(* Logix 5000 project; controller TFF vendor 1 type 14 code 107 rev 33.11; software revision 33.04; part 26 of 38 *)
(* tags used below, declared in another part *)
   Address : DINT;   // Temp Address
   Index : DINT;   // Index
   PCV101_PID_Settings : INT;
   TIME : DINT[2];
   AnalogOutput : AnalogOutput[25];   // Analog Output Array
   AnalogPoint : AnalogInput[50];   // Analog Input Array
   ControlLoop : ControlLoop[20];   // Control Loop Array
   ControlLoop_PCV201 : ALIAS FOR ControlLoop[5];
   ControlLoop_PCV201_5ms : ALIAS FOR ControlLoop[6];
   ControlLoop_PCV201_CV : REAL;   // Control Value
   ControlLoop_PCV201_RAMP_OUT : REAL;   // Ramp Output
   ControlLoop_TIC101 : ALIAS FOR ControlLoop[7];
   ExternalTCU : BOOL;   // Use of External TCU
   LI101 : ALIAS FOR AnalogPoint[44];
   PCV201_Control : PCV_Control;   // PCV201 Control UDT
   Phase0 : ALIAS FOR Phase[0];   // Phase 0
   SysControl : SysControl;   // General system status and command
   Tank : TankManagement;   // Tank Management
   TCU101_AO : ALIAS FOR AnalogOutput[6];
   TCU101ON : ALIAS FOR DigitalOutput[20];
   TIC101Control : TCUControl;
(* Process, continued *)

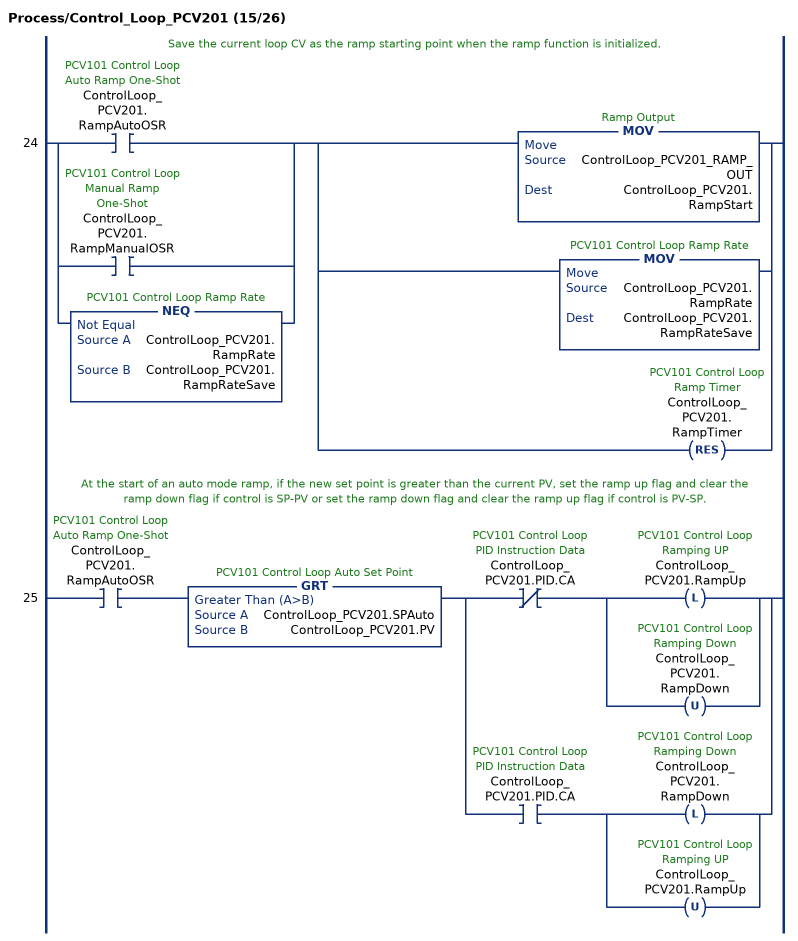
   [picture p239: Process/Control_Loop_PCV201 rungs 24-25]
   // Save the current loop CV as the ramp starting point when the ramp function is initialized.
   24: [XIC(ControlLoop_PCV201.RampAutoOSR) ,XIC(ControlLoop_PCV201.RampManualOSR) ,NEQ(ControlLoop_PCV201.RampRate,ControlLoop_PCV201.RampRateSave) ][MOV(ControlLoop_PCV201_RAMP_OUT,ControlLoop_PCV201.RampStart) ,MOV(ControlLoop_PCV201.RampRate,ControlLoop_PCV201.RampRateSave) ,RES(ControlLoop_PCV201.RampTimer) ];
   // At the start of an auto mode ramp, if the new set point is greater than the current PV, set the ramp up flag and clear the ramp down flag if control is SP-PV or set the ramp down flag and clear the ramp up flag if control is PV-SP.
   25: XIC(ControlLoop_PCV201.RampAutoOSR)GRT(ControlLoop_PCV201.SPAuto,ControlLoop_PCV201.PV)[XIO(ControlLoop_PCV201.PID.CA) [OTL(ControlLoop_PCV201.RampUp) ,OTU(ControlLoop_PCV201.RampDown) ] ,XIC(ControlLoop_PCV201.PID.CA) [OTL(ControlLoop_PCV201.RampDown) ,OTU(ControlLoop_PCV201.RampUp) ] ];
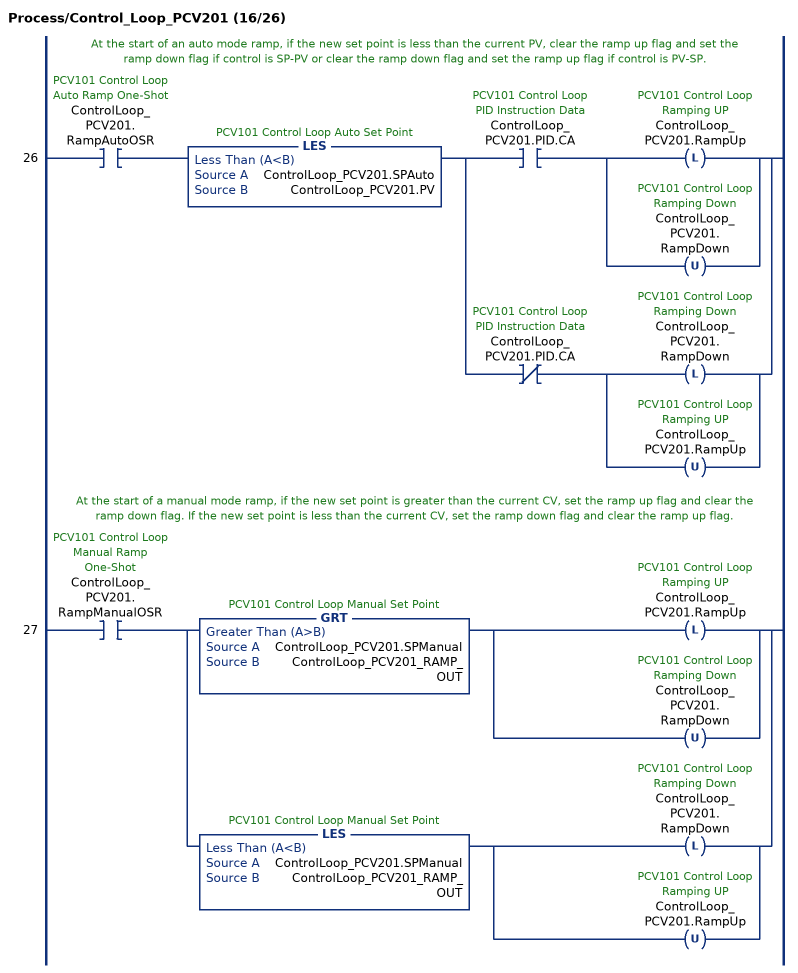
   // At the start of an auto mode ramp, if the new set point is less than the current PV, clear the ramp up flag and set the ramp down flag if control is SP-PV or clear the ramp down flag and set the ramp up flag if control is PV-SP.
   26: XIC(ControlLoop_PCV201.RampAutoOSR)LES(ControlLoop_PCV201.SPAuto,ControlLoop_PCV201.PV)[XIC(ControlLoop_PCV201.PID.CA) [OTL(ControlLoop_PCV201.RampUp) ,OTU(ControlLoop_PCV201.RampDown) ] ,XIO(ControlLoop_PCV201.PID.CA) [OTL(ControlLoop_PCV201.RampDown) ,OTU(ControlLoop_PCV201.RampUp) ] ];
   // At the start of a manual mode ramp, if the new set point is greater than the current CV, set the ramp up flag and clear the ramp down flag. If the new set point is less than the current CV, set the ramp down flag and clear the ramp up flag.
   27: XIC(ControlLoop_PCV201.RampManualOSR)[GRT(ControlLoop_PCV201.SPManual,ControlLoop_PCV201_RAMP_OUT) [OTL(ControlLoop_PCV201.RampUp) ,OTU(ControlLoop_PCV201.RampDown) ] ,LES(ControlLoop_PCV201.SPManual,ControlLoop_PCV201_RAMP_OUT) [OTL(ControlLoop_PCV201.RampDown) ,OTU(ControlLoop_PCV201.RampUp) ] ];
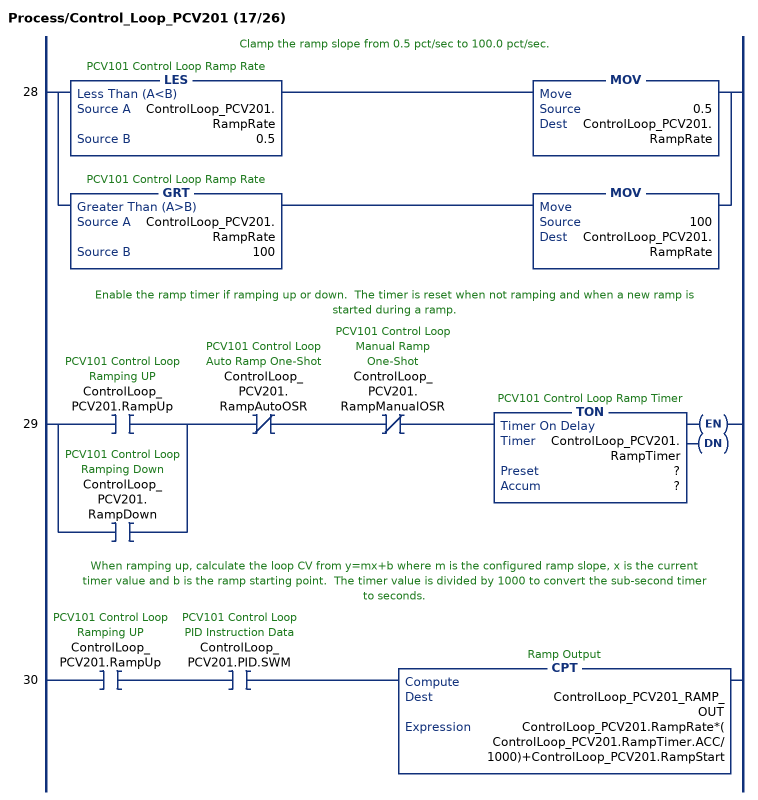
   // Clamp the ramp slope from 0.5 pct/sec to 100.0 pct/sec.
   28: [LES(ControlLoop_PCV201.RampRate,0.5) MOV(0.5,ControlLoop_PCV201.RampRate) ,GRT(ControlLoop_PCV201.RampRate,100) MOV(100,ControlLoop_PCV201.RampRate) ];
   // Enable the ramp timer if ramping up or down.  The timer is reset when not ramping and when a new ramp is started during a ramp.
   29: [XIC(ControlLoop_PCV201.RampUp) ,XIC(ControlLoop_PCV201.RampDown) ]XIO(ControlLoop_PCV201.RampAutoOSR)XIO(ControlLoop_PCV201.RampManualOSR)TON(ControlLoop_PCV201.RampTimer,?,?);
   // When ramping up, calculate the loop CV from y=mx+b where m is the configured ramp slope, x is the current timer value and b is the ramp starting point.  The timer value is divided by 1000 to convert the sub-second timer to seconds.
   30: XIC(ControlLoop_PCV201.RampUp)XIC(ControlLoop_PCV201.PID.SWM)CPT(ControlLoop_PCV201_RAMP_OUT,ControlLoop_PCV201.RampRate*(ControlLoop_PCV201.RampTimer.ACC/1000)+ControlLoop_PCV201.RampStart);
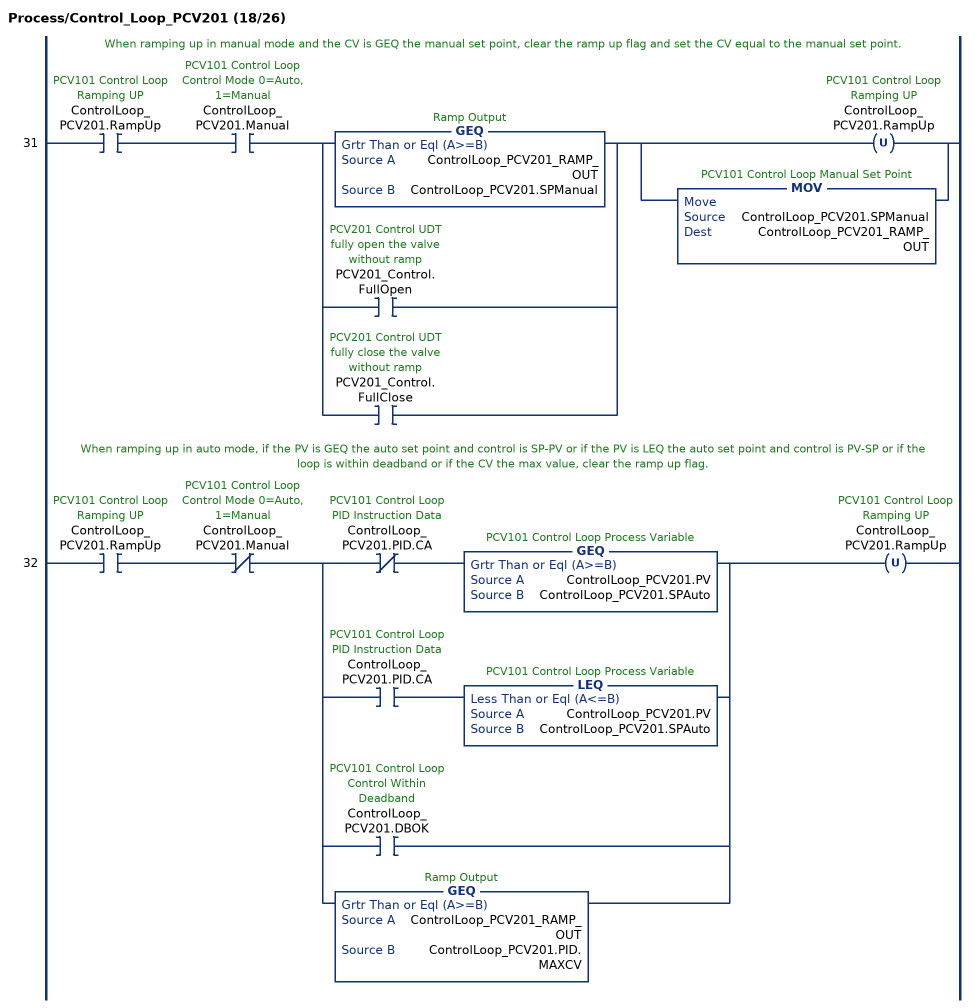
   // When ramping up in manual mode and the CV is GEQ the manual set point, clear the ramp up flag and set the CV equal to the manual set point.
   31: XIC(ControlLoop_PCV201.RampUp)XIC(ControlLoop_PCV201.Manual)[GEQ(ControlLoop_PCV201_RAMP_OUT,ControlLoop_PCV201.SPManual) ,XIC(PCV201_Control.FullOpen) ,XIC(PCV201_Control.FullClose) ][OTU(ControlLoop_PCV201.RampUp) ,MOV(ControlLoop_PCV201.SPManual,ControlLoop_PCV201_RAMP_OUT) ];
   // When ramping up in auto mode, if the PV is GEQ the auto set point and control is SP-PV or if the PV is LEQ the auto set point and control is PV-SP or if the loop is within deadband or if the CV the max value, clear the ramp up flag.
   32: XIC(ControlLoop_PCV201.RampUp)XIO(ControlLoop_PCV201.Manual)[XIO(ControlLoop_PCV201.PID.CA) GEQ(ControlLoop_PCV201.PV,ControlLoop_PCV201.SPAuto) ,XIC(ControlLoop_PCV201.PID.CA) LEQ(ControlLoop_PCV201.PV,ControlLoop_PCV201.SPAuto) ,XIC(ControlLoop_PCV201.DBOK) ,GEQ(ControlLoop_PCV201_RAMP_OUT,ControlLoop_PCV201.PID.MAXCV) ]OTU(ControlLoop_PCV201.RampUp);
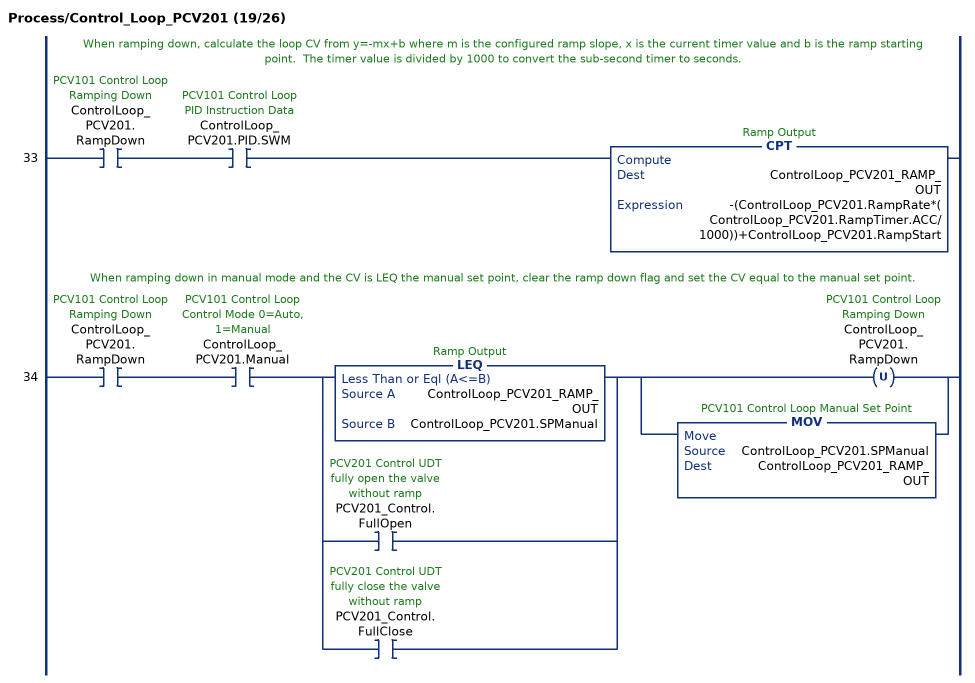
   // When ramping down, calculate the loop CV from y=-mx+b where m is the configured ramp slope, x is the current timer value and b is the ramp starting point.  The timer value is divided by 1000 to convert the sub-second timer to seconds.
   33: XIC(ControlLoop_PCV201.RampDown)XIC(ControlLoop_PCV201.PID.SWM)CPT(ControlLoop_PCV201_RAMP_OUT,-(ControlLoop_PCV201.RampRate*(ControlLoop_PCV201.RampTimer.ACC/1000))+ControlLoop_PCV201.RampStart);
   // When ramping down in manual mode and the CV is LEQ the manual set point, clear the ramp down flag and set the CV equal to the manual set point.
   34: XIC(ControlLoop_PCV201.RampDown)XIC(ControlLoop_PCV201.Manual)[LEQ(ControlLoop_PCV201_RAMP_OUT,ControlLoop_PCV201.SPManual) ,XIC(PCV201_Control.FullOpen) ,XIC(PCV201_Control.FullClose) ][OTU(ControlLoop_PCV201.RampDown) ,MOV(ControlLoop_PCV201.SPManual,ControlLoop_PCV201_RAMP_OUT) ];
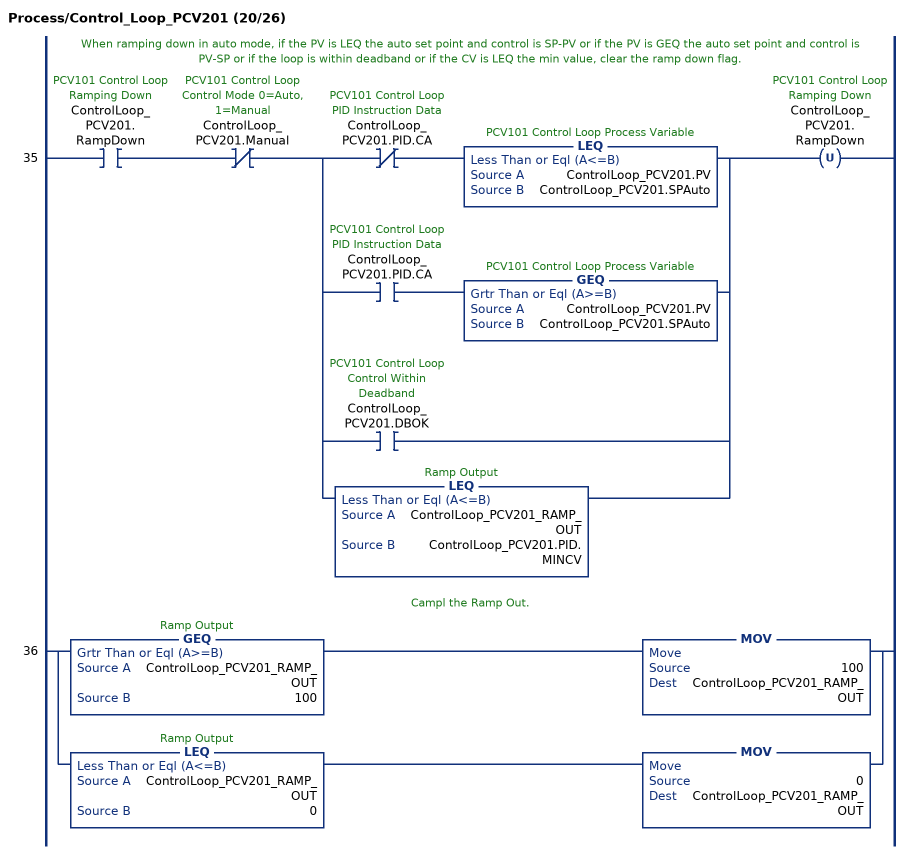
   // When ramping down in auto mode, if the PV is LEQ the auto set point and control is SP-PV or if the PV is GEQ the auto set point and control is PV-SP or if the loop is within deadband or if the CV is LEQ the min value, clear the ramp down flag.
   35: XIC(ControlLoop_PCV201.RampDown)XIO(ControlLoop_PCV201.Manual)[XIO(ControlLoop_PCV201.PID.CA) LEQ(ControlLoop_PCV201.PV,ControlLoop_PCV201.SPAuto) ,XIC(ControlLoop_PCV201.PID.CA) GEQ(ControlLoop_PCV201.PV,ControlLoop_PCV201.SPAuto) ,XIC(ControlLoop_PCV201.DBOK) ,LEQ(ControlLoop_PCV201_RAMP_OUT,ControlLoop_PCV201.PID.MINCV) ]OTU(ControlLoop_PCV201.RampDown);
   // Campl the Ramp Out.
   36: [GEQ(ControlLoop_PCV201_RAMP_OUT,100) MOV(100,ControlLoop_PCV201_RAMP_OUT) ,LEQ(ControlLoop_PCV201_RAMP_OUT,0) MOV(0,ControlLoop_PCV201_RAMP_OUT) ];
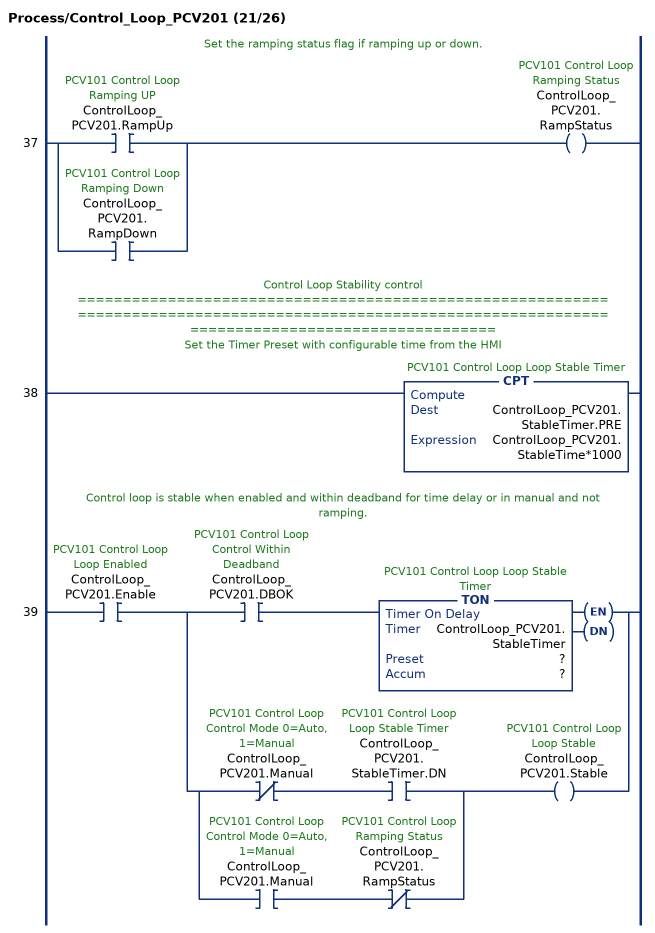
   // Set the ramping status flag if ramping up or down.
   37: [XIC(ControlLoop_PCV201.RampUp) ,XIC(ControlLoop_PCV201.RampDown) ]OTE(ControlLoop_PCV201.RampStatus);
   // Control Loop Stability control
   // ========================================================================================================================================================
   // Set the Timer Preset with configurable time from the HMI
   38: CPT(ControlLoop_PCV201.StableTimer.PRE,ControlLoop_PCV201.StableTime*1000);
   // Control loop is stable when enabled and within deadband for time delay or in manual and not ramping.
   39: XIC(ControlLoop_PCV201.Enable)[XIC(ControlLoop_PCV201.DBOK) TON(ControlLoop_PCV201.StableTimer,?,?) ,[XIO(ControlLoop_PCV201.Manual) XIC(ControlLoop_PCV201.StableTimer.DN) ,XIC(ControlLoop_PCV201.Manual) XIO(ControlLoop_PCV201.RampStatus) ] OTE(ControlLoop_PCV201.Stable) ];
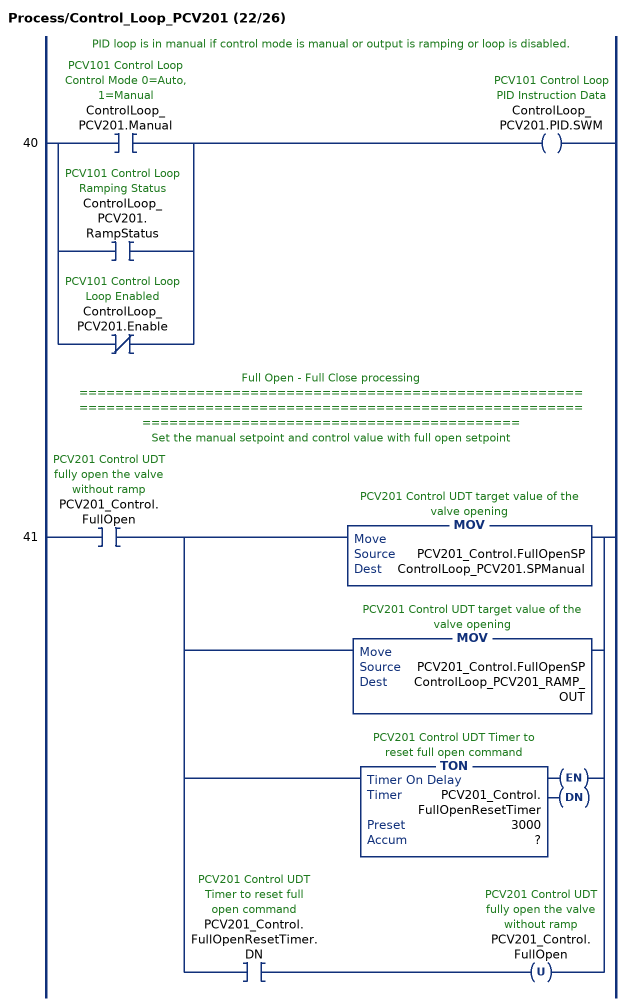
   // PID loop is in manual if control mode is manual or output is ramping or loop is disabled.
   40: [XIC(ControlLoop_PCV201.Manual) ,XIC(ControlLoop_PCV201.RampStatus) ,XIO(ControlLoop_PCV201.Enable) ]OTE(ControlLoop_PCV201.PID.SWM);
   // Full Open - Full Close processing
   // ==========================================================================================================================================================
   // Set the manual setpoint and control value with full open setpoint
   41: XIC(PCV201_Control.FullOpen)[MOV(PCV201_Control.FullOpenSP,ControlLoop_PCV201.SPManual) ,MOV(PCV201_Control.FullOpenSP,ControlLoop_PCV201_RAMP_OUT) ,TON(PCV201_Control.FullOpenResetTimer,?,?) ,XIC(PCV201_Control.FullOpenResetTimer.DN) OTU(PCV201_Control.FullOpen) ];
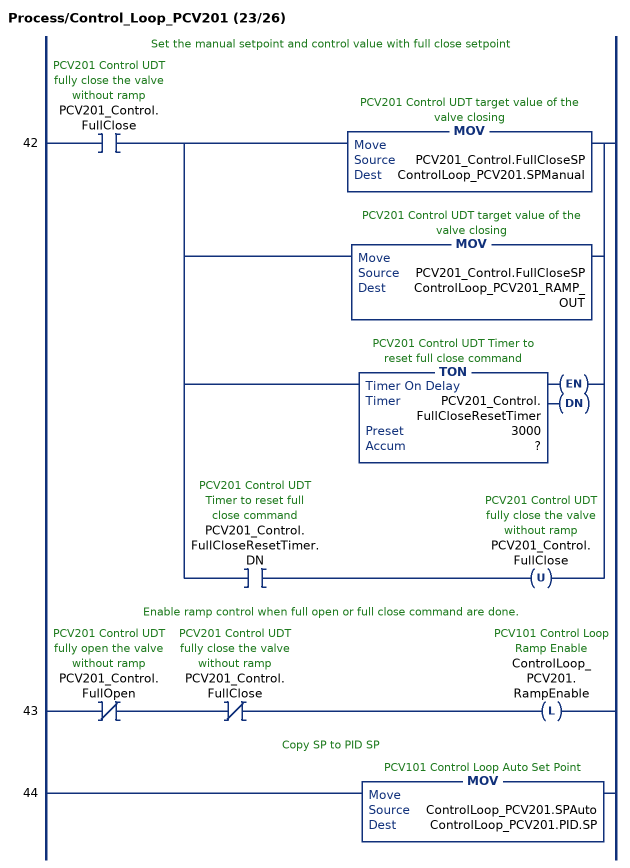
   // Set the manual setpoint and control value with full close setpoint
   42: XIC(PCV201_Control.FullClose)[MOV(PCV201_Control.FullCloseSP,ControlLoop_PCV201.SPManual) ,MOV(PCV201_Control.FullCloseSP,ControlLoop_PCV201_RAMP_OUT) ,TON(PCV201_Control.FullCloseResetTimer,?,?) ,XIC(PCV201_Control.FullCloseResetTimer.DN) OTU(PCV201_Control.FullClose) ];
   // Enable ramp control when full open or full close command are done.
   43: XIO(PCV201_Control.FullOpen)XIO(PCV201_Control.FullClose)OTL(ControlLoop_PCV201.RampEnable);
   // Copy SP to PID SP
   44: MOV(ControlLoop_PCV201.SPAuto,ControlLoop_PCV201.PID.SP);
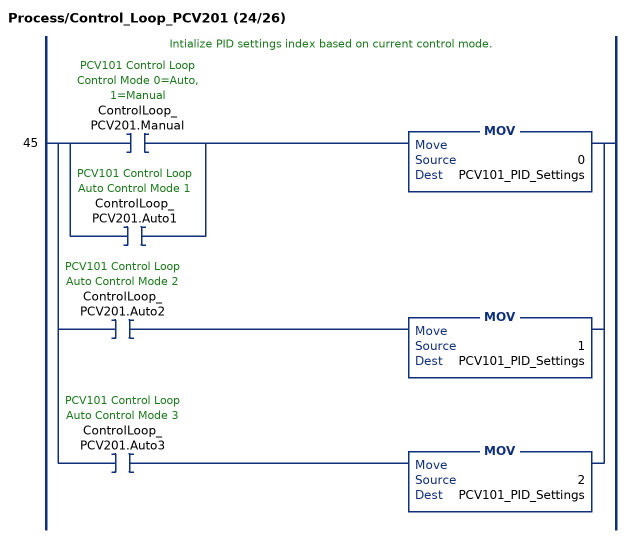
   // Intialize PID settings index based on current control mode.
   45: [[XIC(ControlLoop_PCV201.Manual) ,XIC(ControlLoop_PCV201.Auto1) ] MOV(0,PCV101_PID_Settings) ,XIC(ControlLoop_PCV201.Auto2) MOV(1,PCV101_PID_Settings) ,XIC(ControlLoop_PCV201.Auto3) MOV(2,PCV101_PID_Settings) ];
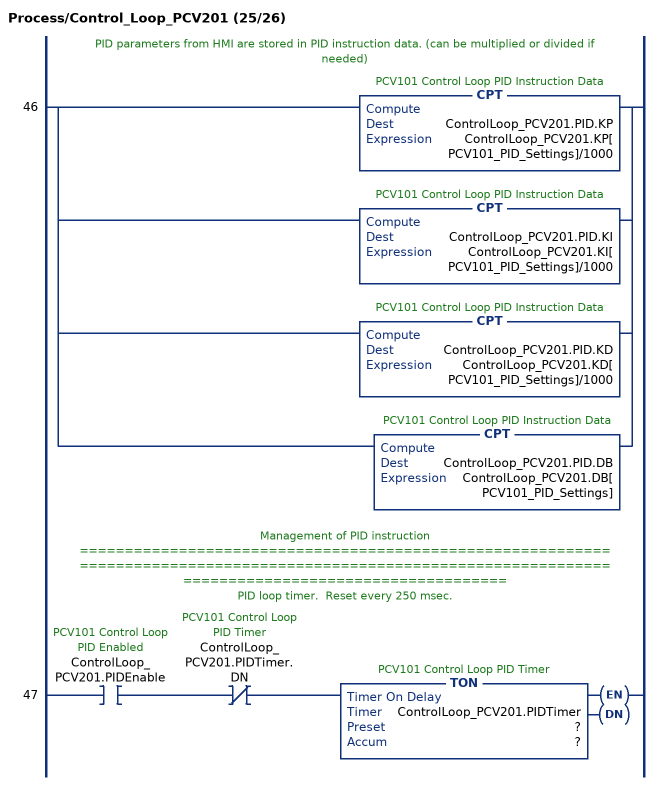
   // PID parameters from HMI are stored in PID instruction data. (can be multiplied or divided if needed)
   46: [CPT(ControlLoop_PCV201.PID.KP,ControlLoop_PCV201.KP[PCV101_PID_Settings]/1000) ,CPT(ControlLoop_PCV201.PID.KI,ControlLoop_PCV201.KI[PCV101_PID_Settings]/1000) ,CPT(ControlLoop_PCV201.PID.KD,ControlLoop_PCV201.KD[PCV101_PID_Settings]/1000) ,CPT(ControlLoop_PCV201.PID.DB,ControlLoop_PCV201.DB[PCV101_PID_Settings]) ];
   // Management of PID instruction
   // ==========================================================================================================================================================
   // PID loop timer.  Reset every 250 msec.
   47: XIC(ControlLoop_PCV201.PIDEnable)XIO(ControlLoop_PCV201.PIDTimer.DN)TON(ControlLoop_PCV201.PIDTimer,?,?);
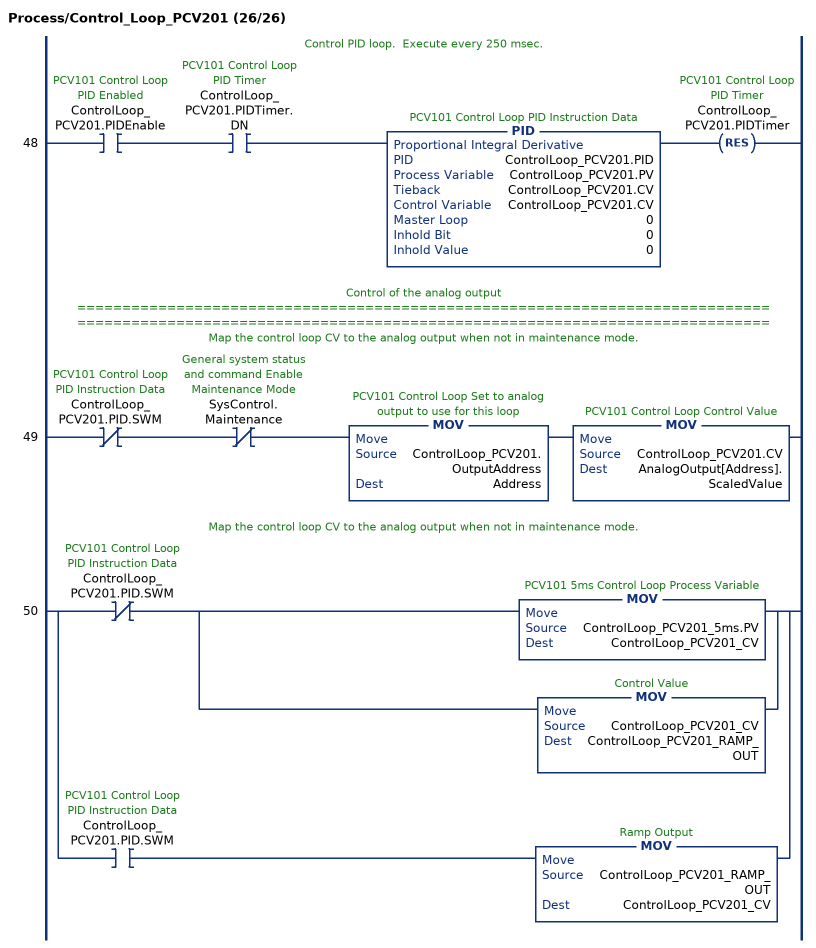
   // Control PID loop.  Execute every 250 msec.
   48: XIC(ControlLoop_PCV201.PIDEnable)XIC(ControlLoop_PCV201.PIDTimer.DN)PID(ControlLoop_PCV201.PID,ControlLoop_PCV201.PV,ControlLoop_PCV201.CV,ControlLoop_PCV201.CV,0,0,0)RES(ControlLoop_PCV201.PIDTimer);
   // Control of the analog output
   // ==========================================================================================================================================================
   // Map the control loop CV to the analog output when not in maintenance mode.
   49: XIO(ControlLoop_PCV201.PID.SWM)XIO(SysControl.Maintenance)MOV(ControlLoop_PCV201.OutputAddress,Address)MOV(ControlLoop_PCV201.CV,AnalogOutput[Address].ScaledValue);
   // Map the control loop CV to the analog output when not in maintenance mode.
   50: [XIO(ControlLoop_PCV201.PID.SWM) [MOV(ControlLoop_PCV201_5ms.PV,ControlLoop_PCV201_CV) ,MOV(ControlLoop_PCV201_CV,ControlLoop_PCV201_RAMP_OUT) ] ,XIC(ControlLoop_PCV201.PID.SWM) MOV(ControlLoop_PCV201_RAMP_OUT,ControlLoop_PCV201_CV) ];
END_ROUTINE

ROUTINE Control_Loop_TIC101   (* ladder *)
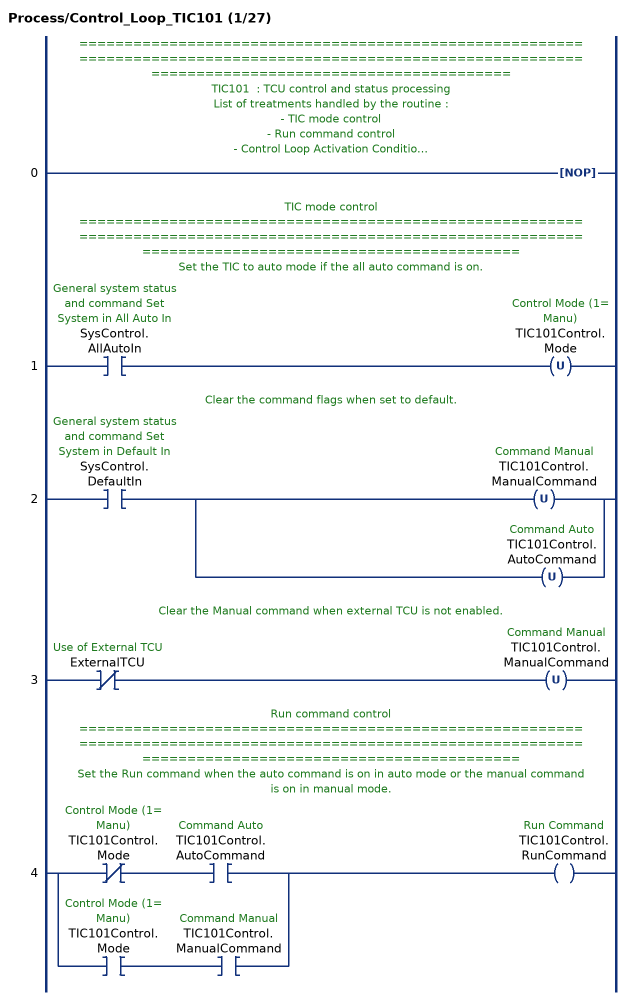
   // ========================================================================================================================================================
   //                                                                                                    TIC101  : TCU control and status processing
   //                                                     List of treatments handled by the routine :
   //                                                     - TIC mode control
   //                                                        - Run command control
   //                                                          - Control Loop Activation Condition
   //                                                          - Control Loop initialization
   //                                                          - Mode control
   //                                                          - Control Loop deadband calculation
   //                                                          - Management of ramping control
   //                                                            - Management of SP Offset
   //                                                          - Control Loop Stability control
   //                                                          - Control Loop manual state control
   //                                                          - Management of PID instruction
   //                                                          - Control of the analog output
   //                                                     -----------------------------------------------------------------------------------------------------------------------------------------------------
   //                                                     History
   // 		2019-DEC-24 - Merck - Q. Spindler - Initial version for Candidate Release 1.00.00.00.a
   // 		2020-SEP-09 - Merck - Q. Spindler - Modifications for Candidate Release 1.00.00.00.d
   // 					- Add ControlLoop Enable and not manual condition for DBOK status
   // 				   	- Clear Manual command when ExternalTCU is disabled
   // 		2021-APR-16 - Merck - Q. Spindler - Modifications for Candidate Release 1.00.00.00.e
   //                                        - Add Initialize address if no mode selected.
   //                       - Change TIC Output Range to 50
   // ========================================================================================================================================================
   0: NOP();
   // TIC mode control
   // ==========================================================================================================================================================
   // Set the TIC to auto mode if the all auto command is on.
   1: XIC(SysControl.AllAutoIn)OTU(TIC101Control.Mode);
   // Clear the command flags when set to default.
   2: XIC(SysControl.DefaultIn)[OTU(TIC101Control.ManualCommand) ,OTU(TIC101Control.AutoCommand) ];
   // Clear the Manual command when external TCU is not enabled.
   3: XIO(ExternalTCU)OTU(TIC101Control.ManualCommand);
   // Run command control
   // ==========================================================================================================================================================
   // Set the Run command when the auto command is on in auto mode or the manual command is on in manual mode.
   4: [XIO(TIC101Control.Mode) XIC(TIC101Control.AutoCommand) ,XIC(TIC101Control.Mode) XIC(TIC101Control.ManualCommand) ]OTE(TIC101Control.RunCommand);
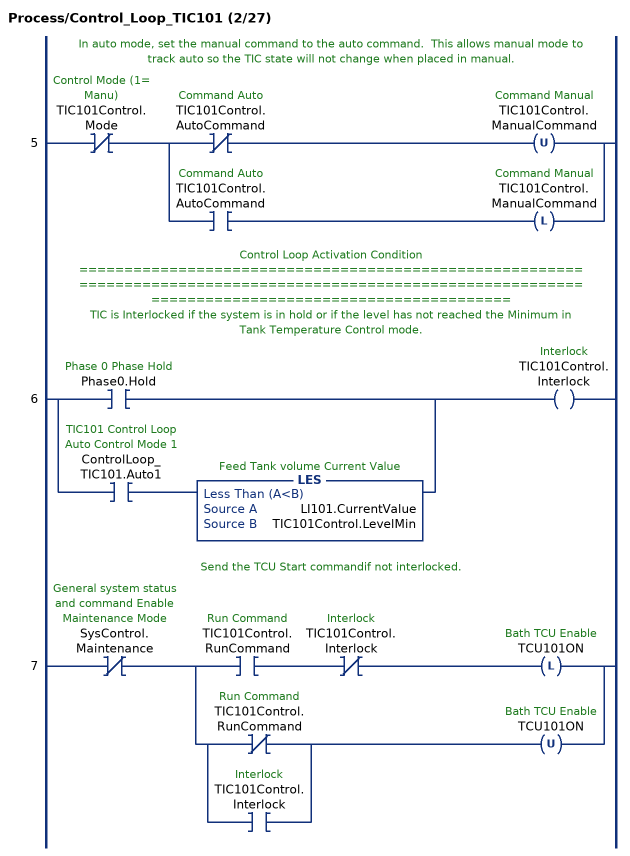
   // In auto mode, set the manual command to the auto command.  This allows manual mode to track auto so the TIC state will not change when placed in manual.
   5: XIO(TIC101Control.Mode)[XIO(TIC101Control.AutoCommand) OTU(TIC101Control.ManualCommand) ,XIC(TIC101Control.AutoCommand) OTL(TIC101Control.ManualCommand) ];
   // Control Loop Activation Condition
   // ========================================================================================================================================================
   // TIC is Interlocked if the system is in hold or if the level has not reached the Minimum in Tank Temperature Control mode.
   6: [XIC(Phase0.Hold) ,XIC(ControlLoop_TIC101.Auto1) LES(LI101.CurrentValue,TIC101Control.LevelMin) ]OTE(TIC101Control.Interlock);
   // Send the TCU Start commandif not interlocked.
   7: XIO(SysControl.Maintenance)[XIC(TIC101Control.RunCommand) XIO(TIC101Control.Interlock) OTL(TCU101ON) ,[XIO(TIC101Control.RunCommand) ,XIC(TIC101Control.Interlock) ] OTU(TCU101ON) ];
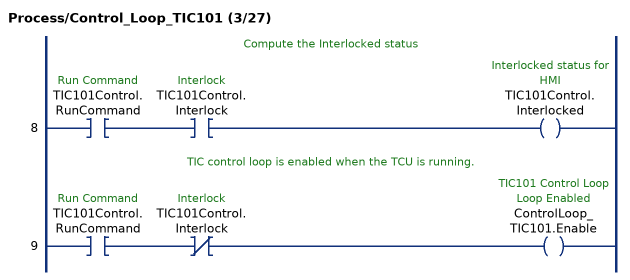
   // Compute the Interlocked status
   8: XIC(TIC101Control.RunCommand)XIC(TIC101Control.Interlock)OTE(TIC101Control.Interlocked);
   // TIC control loop is enabled when the TCU is running.
   9: XIC(TIC101Control.RunCommand)XIO(TIC101Control.Interlock)OTE(ControlLoop_TIC101.Enable);
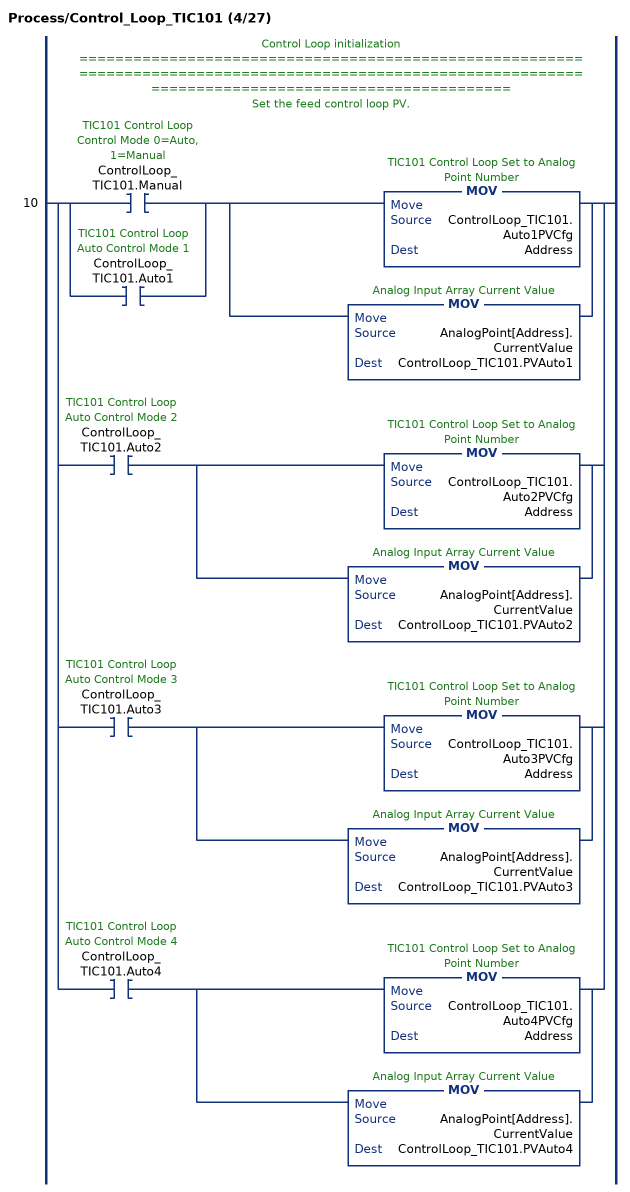
   // Control Loop initialization
   // ========================================================================================================================================================
   // Set the feed control loop PV.
   10: [[[XIC(ControlLoop_TIC101.Manual) ,XIC(ControlLoop_TIC101.Auto1) ] [MOV(ControlLoop_TIC101.Auto1PVCfg,Address) ,MOV(AnalogPoint[Address].CurrentValue,ControlLoop_TIC101.PVAuto1) ] ,XIC(ControlLoop_TIC101.Auto2) [MOV(ControlLoop_TIC101.Auto2PVCfg,Address) ,MOV(AnalogPoint[Address].CurrentValue,ControlLoop_TIC101.PVAuto2) ] ] ,XIC(ControlLoop_TIC101.Auto3) [MOV(ControlLoop_TIC101.Auto3PVCfg,Address) ,MOV(AnalogPoint[Address].CurrentValue,ControlLoop_TIC101.PVAuto3) ] ,XIC(ControlLoop_TIC101.Auto4) [MOV(ControlLoop_TIC101.Auto4PVCfg,Address) ,MOV(AnalogPoint[Address].CurrentValue,ControlLoop_TIC101.PVAuto4) ] ];
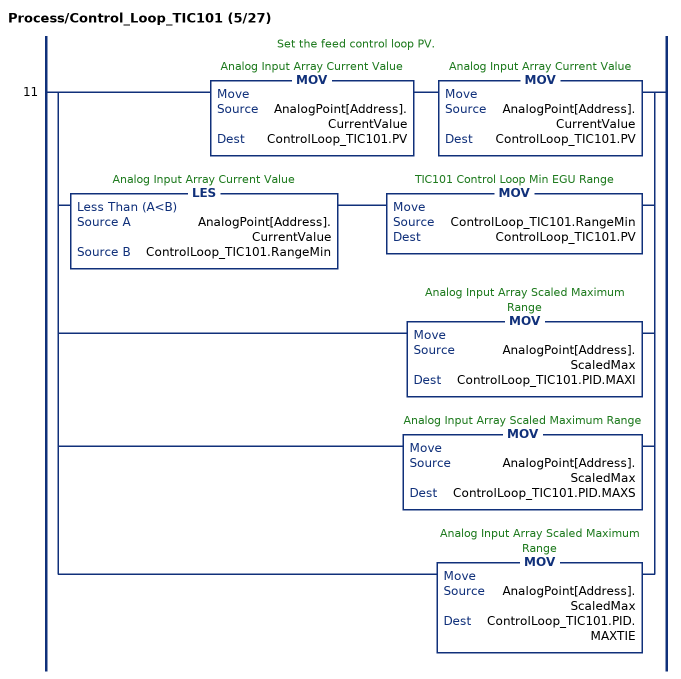
   // Set the feed control loop PV.
   11: [MOV(AnalogPoint[Address].CurrentValue,ControlLoop_TIC101.PV) MOV(AnalogPoint[Address].CurrentValue,ControlLoop_TIC101.PV) ,LES(AnalogPoint[Address].CurrentValue,ControlLoop_TIC101.RangeMin) MOV(ControlLoop_TIC101.RangeMin,ControlLoop_TIC101.PV) ,MOV(AnalogPoint[Address].ScaledMax,ControlLoop_TIC101.PID.MAXI) ,MOV(AnalogPoint[Address].ScaledMax,ControlLoop_TIC101.PID.MAXS) ,MOV(AnalogPoint[Address].ScaledMax,ControlLoop_TIC101.PID.MAXTIE) ];
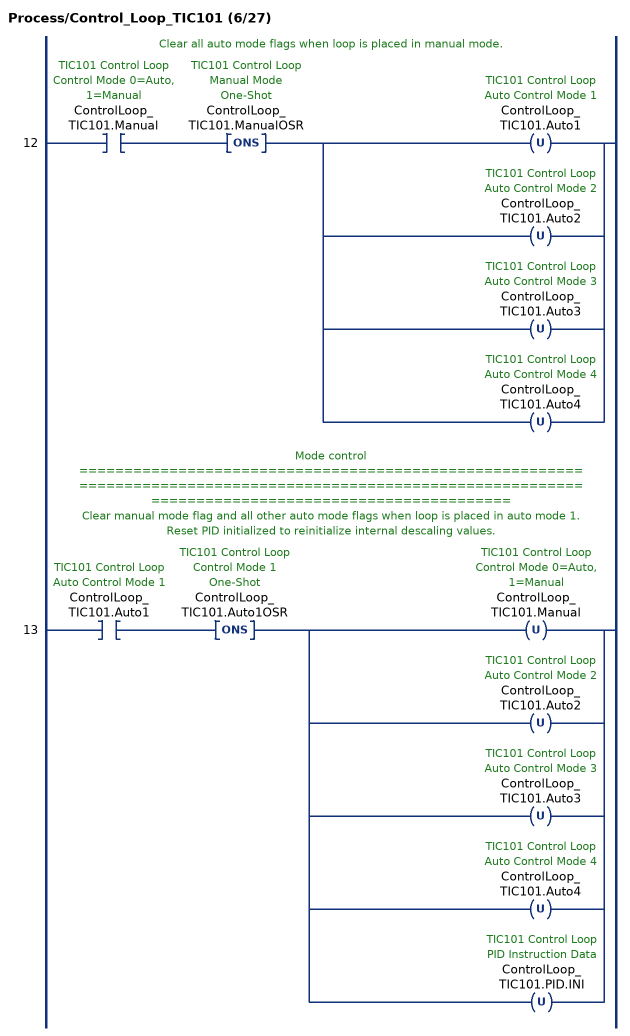
   // Clear all auto mode flags when loop is placed in manual mode.
   12: XIC(ControlLoop_TIC101.Manual)ONS(ControlLoop_TIC101.ManualOSR)[OTU(ControlLoop_TIC101.Auto1) ,OTU(ControlLoop_TIC101.Auto2) ,OTU(ControlLoop_TIC101.Auto3) ,OTU(ControlLoop_TIC101.Auto4) ];
   // Mode control
   // ========================================================================================================================================================
   // Clear manual mode flag and all other auto mode flags when loop is placed in auto mode 1. Reset PID initialized to reinitialize internal descaling values.
   13: XIC(ControlLoop_TIC101.Auto1)ONS(ControlLoop_TIC101.Auto1OSR)[OTU(ControlLoop_TIC101.Manual) ,OTU(ControlLoop_TIC101.Auto2) ,OTU(ControlLoop_TIC101.Auto3) ,OTU(ControlLoop_TIC101.Auto4) ,OTU(ControlLoop_TIC101.PID.INI) ];
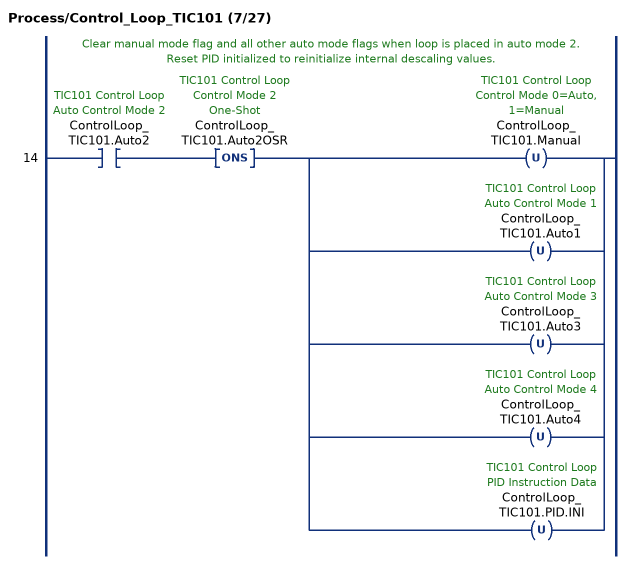
   // Clear manual mode flag and all other auto mode flags when loop is placed in auto mode 2. Reset PID initialized to reinitialize internal descaling values.
   14: XIC(ControlLoop_TIC101.Auto2)ONS(ControlLoop_TIC101.Auto2OSR)[OTU(ControlLoop_TIC101.Manual) ,OTU(ControlLoop_TIC101.Auto1) ,OTU(ControlLoop_TIC101.Auto3) ,OTU(ControlLoop_TIC101.Auto4) ,OTU(ControlLoop_TIC101.PID.INI) ];
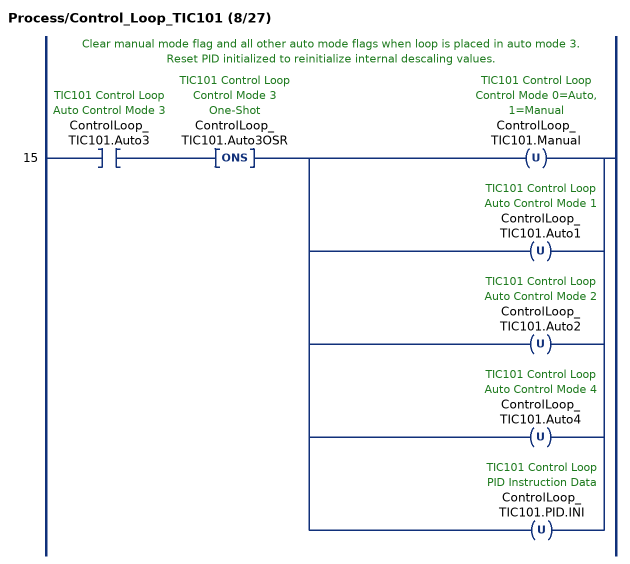
   // Clear manual mode flag and all other auto mode flags when loop is placed in auto mode 3. Reset PID initialized to reinitialize internal descaling values.
   15: XIC(ControlLoop_TIC101.Auto3)ONS(ControlLoop_TIC101.Auto3OSR)[OTU(ControlLoop_TIC101.Manual) ,OTU(ControlLoop_TIC101.Auto1) ,OTU(ControlLoop_TIC101.Auto2) ,OTU(ControlLoop_TIC101.Auto4) ,OTU(ControlLoop_TIC101.PID.INI) ];
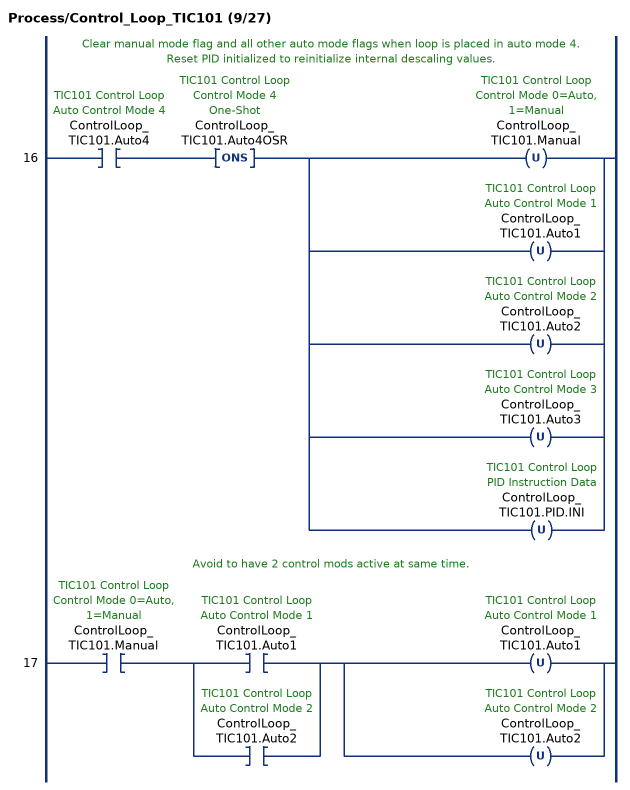
   // Clear manual mode flag and all other auto mode flags when loop is placed in auto mode 4. Reset PID initialized to reinitialize internal descaling values.
   16: XIC(ControlLoop_TIC101.Auto4)ONS(ControlLoop_TIC101.Auto4OSR)[OTU(ControlLoop_TIC101.Manual) ,OTU(ControlLoop_TIC101.Auto1) ,OTU(ControlLoop_TIC101.Auto2) ,OTU(ControlLoop_TIC101.Auto3) ,OTU(ControlLoop_TIC101.PID.INI) ];
   // Avoid to have 2 control mods active at same time.
   17: XIC(ControlLoop_TIC101.Manual)[XIC(ControlLoop_TIC101.Auto1) ,XIC(ControlLoop_TIC101.Auto2) ][OTU(ControlLoop_TIC101.Auto1) ,OTU(ControlLoop_TIC101.Auto2) ];
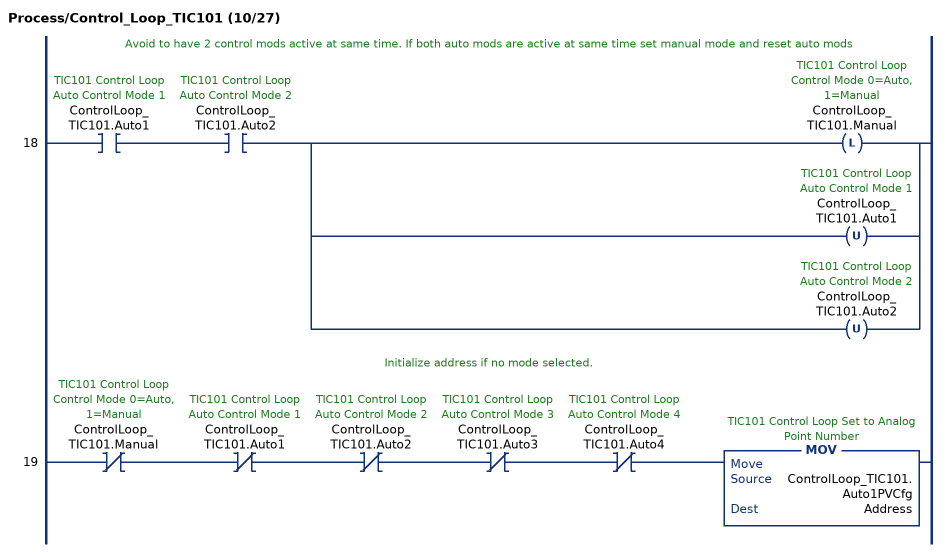
   // Avoid to have 2 control mods active at same time. If both auto mods are active at same time set manual mode and reset auto mods
   18: XIC(ControlLoop_TIC101.Auto1)XIC(ControlLoop_TIC101.Auto2)[OTL(ControlLoop_TIC101.Manual) ,OTU(ControlLoop_TIC101.Auto1) ,OTU(ControlLoop_TIC101.Auto2) ];
   // Initialize address if no mode selected.
   19: XIO(ControlLoop_TIC101.Manual)XIO(ControlLoop_TIC101.Auto1)XIO(ControlLoop_TIC101.Auto2)XIO(ControlLoop_TIC101.Auto3)XIO(ControlLoop_TIC101.Auto4)MOV(ControlLoop_TIC101.Auto1PVCfg,Address);
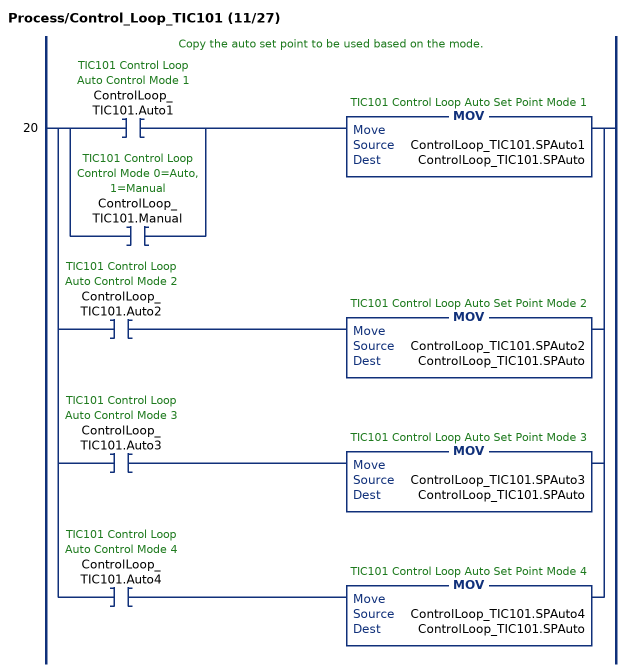
   // Copy the auto set point to be used based on the mode.
   20: [[XIC(ControlLoop_TIC101.Auto1) ,XIC(ControlLoop_TIC101.Manual) ] MOV(ControlLoop_TIC101.SPAuto1,ControlLoop_TIC101.SPAuto) ,XIC(ControlLoop_TIC101.Auto2) MOV(ControlLoop_TIC101.SPAuto2,ControlLoop_TIC101.SPAuto) ,XIC(ControlLoop_TIC101.Auto3) MOV(ControlLoop_TIC101.SPAuto3,ControlLoop_TIC101.SPAuto) ,XIC(ControlLoop_TIC101.Auto4) MOV(ControlLoop_TIC101.SPAuto4,ControlLoop_TIC101.SPAuto) ];
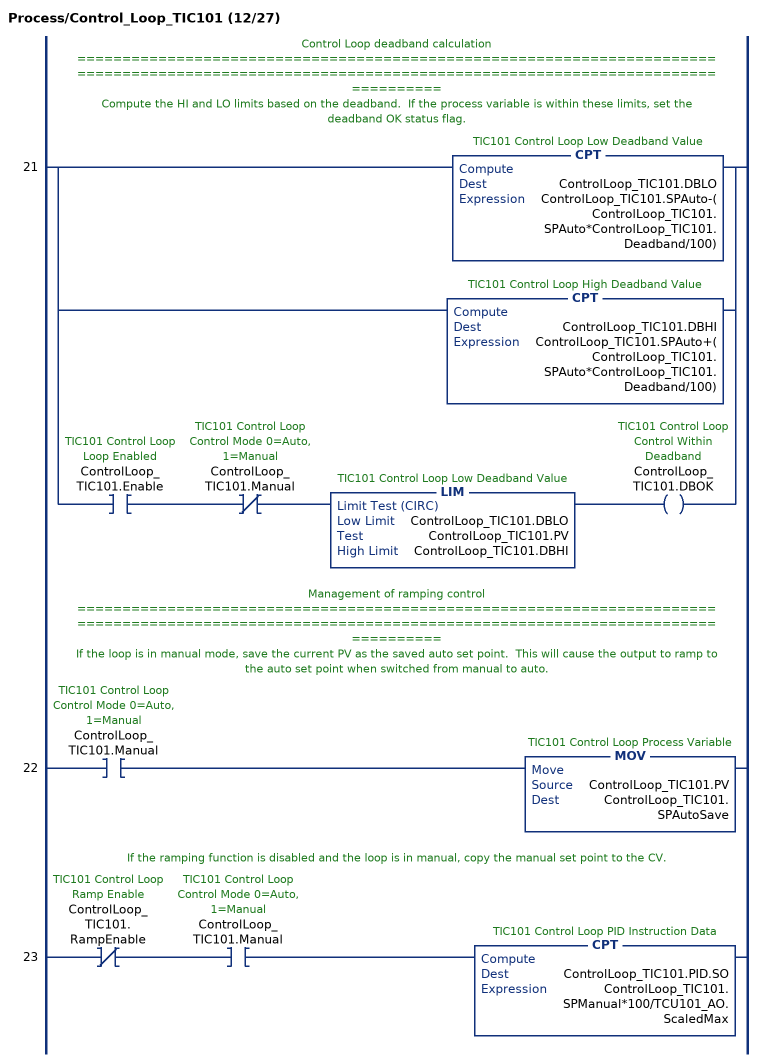
   // Control Loop deadband calculation
   // ========================================================================================================================================================
   // Compute the HI and LO limits based on the deadband.  If the process variable is within these limits, set the deadband OK status flag.
   21: [CPT(ControlLoop_TIC101.DBLO,ControlLoop_TIC101.SPAuto-(ControlLoop_TIC101.SPAuto*ControlLoop_TIC101.Deadband/100)) ,CPT(ControlLoop_TIC101.DBHI,ControlLoop_TIC101.SPAuto+(ControlLoop_TIC101.SPAuto*ControlLoop_TIC101.Deadband/100)) ,XIC(ControlLoop_TIC101.Enable) XIO(ControlLoop_TIC101.Manual) LIM(ControlLoop_TIC101.DBLO,ControlLoop_TIC101.PV,ControlLoop_TIC101.DBHI) OTE(ControlLoop_TIC101.DBOK) ];
   // Management of ramping control
   // ========================================================================================================================================================
   // If the loop is in manual mode, save the current PV as the saved auto set point.  This will cause the output to ramp to the auto set point when switched from manual to auto.
   22: XIC(ControlLoop_TIC101.Manual)MOV(ControlLoop_TIC101.PV,ControlLoop_TIC101.SPAutoSave);
   // If the ramping function is disabled and the loop is in manual, copy the manual set point to the CV.
   23: XIO(ControlLoop_TIC101.RampEnable)XIC(ControlLoop_TIC101.Manual)CPT(ControlLoop_TIC101.PID.SO,ControlLoop_TIC101.SPManual*100/TCU101_AO.ScaledMax);
